{attribute 'qualified_only'}
VAR_GLOBAL
	//Input
	StartButton		:	BOOL;
	StopButton		:	BOOL;
	EmergencyStop	:	BOOL;
	Reset			:	BOOL;
	
	SensorEntry		:	BOOL;
	SensorExit		:	BOOL;
	AutoMode		:	BOOL;
	
	
	//Output
	Motor			:	BOOL;
	MotorStopped 	: 	BOOL;
	GreenLamp 		:	BOOL;
	RedLamp 		:	BOOL;
	
	FaultLamp		:	BOOL;
	
	FaultCode 		: 	E_FaultCode;
	
	FaultText : STRING(50) := 'NO FAULT';
	ModeText  : STRING(50) ;
	
	
	Mode : E_ConveyorMode := E_ConveyorMode.AUTO;
	
	
	
	
END_VAR

(* stored: Version 1.1.0.1, ProductVersion 3.1.4026.21
   GVL GVL_IO: Id {4baea8d6-b063-491a-b9b5-ad5ff0cbac32} *)
